(* PLC project Vn_member_read, Beckhoff Automation GmbH TwinCAT PLC Control 3.5.13.21 *)
(* stored: creationDateTime 1970-01-01T00:00:00 *)

PROGRAM Vn_member_read

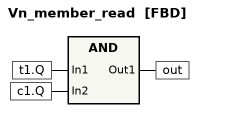
(* FBD diagram, written out as Structured Text *)
out := t1.Q AND c1.Q;
END_PROGRAM
